FUNCTION F_ModR : REAL
(*
Modulo function for real numbers (dividend mod divisor).

Constructor: 		Patryk Panylo
Company:		E. Riexinger GmbH
Date:			20.01.2014
Version:			1.00

Date:			Revision:		Who:				Comment
dd.mm.yyyy		x.xx			Initials			comment

*)
VAR_INPUT
	rDividend						:REAL;
	rDivisor							:REAL := 1.0;
END_VAR
VAR
END_VAR


F_ModR := rDivisor;

IF rDivisor <> 0.0 
THEN
	F_ModR := rDividend - DINT_TO_REAL(F_FloorDN(rDividend / rDivisor)) * rDivisor;
END_IF;

END_FUNCTION

(* stored: Version 1.1.0.1, ProductVersion 3.1.4024.15
   POU F_ModR: Id {f0451ca7-5d22-4d76-9b4b-4586b4a31324}, SpecialFunc None *)
